// TIA Portal V21 export
// export: Created 2026-11-21T13:24:04.7324209Z, ExportSetting WithDefaults, DisplayName Totally Integrated Automation Portal, DisplayVersion V21, DisplayName STEP 7 Professional, DisplayVersion V21, DisplayName STEP 7 Safety, DisplayVersion V21, DisplayName Tech WebApplication, DisplayVersion V21, DisplayName WinCC Basic/Comfort/Advanced, DisplayVersion V21, DisplayName WinCC Unified, DisplayVersion V21
FUNCTION_BLOCK "GuardSafety"   // FB4, F_FBD
{ S7_Optimized_Access := 'TRUE' }
VERSION : 0.1
// Main safety block of the guard's F-runtime group.
// stored: AutoNumber true, IsIECCheckEnabled false, UDAEnableTagReadback false
   VAR
      guard : "Guard";
      hornOn : Bool;
   END_VAR
BEGIN

REGION Network 1: Guard
   // The horn is on while the guard is open.
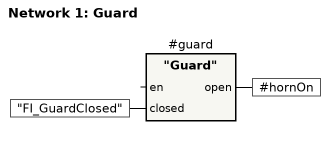
   #guard(closed := "FI_GuardClosed", open => #hornOn);   // "Guard"
END_REGION
END_FUNCTION_BLOCK
